TYPE ET_LoadFromFile_1 :
(
	ET_LoadFromFile_eWaitExecute := 0,
	ET_LoadFromFile_eFileName,
	ET_LoadFromFile_eChkFileExist,
	ET_LoadFromFile_eFileOpen,
	ET_LoadFromFile_eChkFileOpen,
	ET_LoadFromFile_eReadData,
	ET_LoadFromFile_eChkReadData,
	ET_LoadFromFile_eFileClose,
	ET_LoadFromFile_eChkFileClose,
	ET_LoadFromFile_eDone := 197,
	ET_LoadFromFile_eError := 198,
	ET_LoadFromFile_eNoExecute := 199
);
END_TYPE

(* stored: Version 1.1.0.1, ProductVersion 3.1.4024.15
   DUT ET_LoadFromFile_1: Id {695eb735-e5be-43ce-8eff-1419e26447a1} *)
